TYPE ST_TankHMI :
STRUCT
    // ---- Commands (HMI -> PLC) ----
    bAutoMode      : BOOL;
    bStart         : BOOL;
    bStop          : BOOL;
    bReset         : BOOL;
    bPB_ValveIn    : BOOL;
    bPB_ValveOut   : BOOL;
    bPB_Pump       : BOOL;

    // ---- Status (PLC -> HMI) ----
    bLampValveIn   : BOOL;
    bLampValveOut  : BOOL;
    bLampPump      : BOOL;
    bLampHigh      : BOOL;
    bLampLow       : BOOL;
    bFaultActive   : BOOL;
    eState         : E_TankState;
    eFaultCode     : E_TankFault;
	
	rLevel         : REAL; 
END_STRUCT
END_TYPE

(* stored: Version 1.1.0.1
   DUT ST_TankHMI: Id {56d26f25-9aac-45e8-97cf-a41d3db88d3d} *)
